PROGRAM MAIN
VAR
	
	PlcFirstCycle : BOOL := TRUE;
	
	// SHUTTERS
	
	ShutterR1CmdEvent : stShutterCmdEvent;

END_VAR
VAR CONSTANT
	ShutterCleanCmdEvent : stShutterCmdEvent := (
        Execute := FALSE,
        Cmd := ( CommandType := eShutterCmdType.NONE, Position := (Height := 0, Angle := 0 ) ) );
END_VAR


IF PlcFirstCycle THEN
	// Place for code done in first plc cycle
	
	PlcFirstCycle := FALSE;
END_IF


// ------ Run Switches ------
gvlSwitches.SwitchR1Open();
gvlSwitches.SwitchR1Close();


// ------ Run Switche Controllers ------
gvlSwitches.SwitchR1OpenCtrl();
gvlSwitches.SwitchR1CloseCtrl();

// Clear Shutter Commands
ShutterR1CmdEvent := ShutterCleanCmdEvent;

// ------ Run Shutter Commands from Auto sources ------

IF gvlHA.Shutter1EveningScheduleSet THEN
	gvlScheduler.Shutter1EveningScheduler.SetConfig(gvlHA.Shutter1EveningScheduleConfig);
	gvlHA.Shutter1EveningScheduleSet := FALSE;
END_IF



// ------ Run Shutter Commands from Switches ------
gvlShutters.ShutterR1Switch.Process(CmdEvent := ShutterR1CmdEvent);

// ------ Run Shutter Commands from Safety sources ------

// ------ Run Shutter Controllers ------
gvlShutters.ShutterR1Ctrl();

// ------ Run Shutter Actuators ------
gvlShutters.ShutterR1Act();

END_PROGRAM

(* stored: Version 1.1.0.1
   POU MAIN: Id {b477ade9-5e41-44da-827a-03687596879d}, SpecialFunc None *)
